// TIA Portal V21 export
// export: Created 2026-11-10T07:35:05.3480123Z, ExportSetting WithDefaults, DisplayName Totally Integrated Automation Portal, DisplayVersion V21 Update 3, DisplayName STEP 7 Professional, DisplayVersion V21 Update 3, DisplayName STEP 7 Safety, DisplayVersion V21, DisplayName Tech WebApplication, DisplayVersion V21, DisplayName WinCC Basic/Comfort/Advanced, DisplayVersion V21 Update 3, DisplayName WinCC Unified, DisplayVersion V21 Update 3
FUNCTION_BLOCK "FB_Lad_ex045"   // FB90, LAD
{ S7_Optimized_Access := 'TRUE' }
VERSION : 0.1
// stored: AutoNumber true, IsIECCheckEnabled false, IsRetainMemResEnabled false, MemoryReserve 100, SetENOAutomatically false, UDAEnableTagReadback false
   VAR_INPUT
      v_req : Bool;
      v_id : HW_IO;
      v_index : DInt;
      v_mlen : UInt;
   END_VAR
   VAR_OUTPUT
      v_valid : Bool;
      v_busy : Bool;
      v_error : Bool;
      v_status : DWord;
      v_len : UInt;
   END_VAR
   VAR_IN_OUT
      v_record : Array[0..99] of Byte;
   END_VAR
   VAR
      inst { S7_SetPoint := 'True'} : RDREC;
   END_VAR
BEGIN

REGION Network 1: RDREC - Read data record
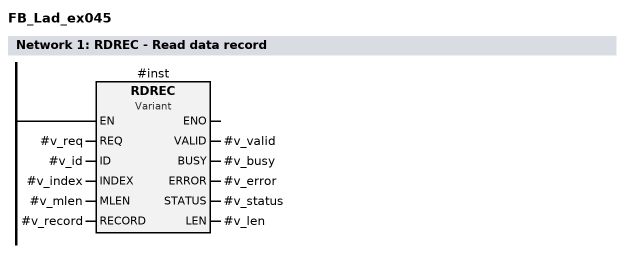
   RUNG wire#powerrail
      { S7_Templates := "[ptr_type := Variant, id_type := HW_IO, index_type := DInt, len_type := UInt]" } #inst.RDREC(REQ := #v_req, ID := #v_id, INDEX := #v_index, MLEN := #v_mlen, VALID => #v_valid, BUSY => #v_busy, ERROR => #v_error, STATUS => #v_status, LEN => #v_len, RECORD := #v_record)
   END_RUNG
   // the same network as SCL:
   #inst(REQ := #v_req,   // RDREC
         ID := #v_id,
         INDEX := #v_index,
         MLEN := #v_mlen,
         RECORD := #v_record,
         VALID => #v_valid,
         BUSY => #v_busy,
         ERROR => #v_error,
         STATUS => #v_status,
         LEN => #v_len);
END_REGION
END_FUNCTION_BLOCK
